(* IEC 61131-3 sources: plc-iiot-stack/src/DUTs/Json, 3 files *)

(* ---- E_JsonError.dut.st ---- *)
// Назначение: причина отказа разбора JSON (FB_JsonFlatParser).
// Документ:   docs/plc_mqtt.md
{attribute 'qualified_only'}
{attribute 'strict'}
TYPE E_JsonError :
(
    None := 0,   // ошибок нет
    Empty := 1,   // пустой вход
    Syntax := 2,   // нарушен синтаксис JSON
    Nested := 3,   // вложенный объект или массив: не поддерживается
    Duplicate := 4,   // ключ повторяется
    TooManyFields := 5,   // полей больше JSON_MAX_FIELDS
    KeyTooLong := 6,   // ключ длиннее JSON_KEY_LEN
    ValueTooLong := 7,   // строка длиннее JSON_STR_LEN
    BadEscape := 8,   // неизвестная escape-последовательность или код вне ASCII
    BadNumber := 9,   // число не по грамматике JSON или вне диапазона REAL
    Trailing := 10   // лишние символы после объекта
) INT;
END_TYPE

(* ---- E_JsonType.dut.st ---- *)
// Назначение: тип значения поля разобранного объекта JSON.
// Документ:   docs/plc_mqtt.md
{attribute 'qualified_only'}
{attribute 'strict'}
TYPE E_JsonType :
(
    Missing := 0,   // поля нет
    Text := 1,   // строка
    Number := 2,   // число
    Boolean := 3,   // true или false
    NullValue := 4   // null
) INT;
END_TYPE

(* ---- ST_JsonField.dut.st ---- *)
// Назначение: поле разобранного плоского объекта JSON.
// Документ:   docs/plc_mqtt.md
{attribute 'qualified_only'}
TYPE ST_JsonField :
STRUCT
    sKey : STRING(GVL_Const.JSON_KEY_LEN);
    eType : E_JsonType := E_JsonType.Missing;
    sText : STRING(GVL_Const.JSON_STR_LEN);   // eType = Text
    lrNumber : LREAL;                         // eType = Number
    xInteger : BOOL;                          // число записано без дробной части и порядка
    xBool : BOOL;                             // eType = Boolean
END_STRUCT
END_TYPE
